(* IEC 61131-3 sources: plc-st-coding-agent/progress/evidence/full_r8_20261110b/native_evidence/codex_minimax-m27/public-easy-04/1, 1 file *)

(* ---- candidate.st ---- *)
FUNCTION_BLOCK FB
VAR_INPUT
    VISCOSITY_OK      : BOOL;
    PASTE_E_STOP_NC   : BOOL;
    DebounceMs        : DINT;
    CycleMs           : DINT;
END_VAR
VAR_OUTPUT
    VFD_RUN           : BOOL;
    PUMP_MAINT_DUE    : BOOL;
    PUMP_RUNTIME_ACC  : LINT;
END_VAR
VAR
    valid_duration     : DINT;
    prev_viscosity_ok  : BOOL;
    prev_paste_e_stop_nc : BOOL;
    prev_valid_duration : DINT;
    prev_vfd_run       : BOOL;
END_VAR

    IF NOT (PASTE_E_STOP_NC AND VISCOSITY_OK) THEN
        VFD_RUN := FALSE;
        valid_duration := 0;
    ELSE
        IF NOT prev_viscosity_ok OR NOT prev_paste_e_stop_nc THEN
            valid_duration := prev_valid_duration + CycleMs;
            VFD_RUN := (valid_duration >= DebounceMs);
        ELSIF prev_vfd_run THEN
            valid_duration := valid_duration + CycleMs;
            VFD_RUN := TRUE;
        ELSE
            valid_duration := valid_duration + CycleMs;
            VFD_RUN := (valid_duration >= DebounceMs);
        END_IF
    END_IF

    IF VFD_RUN THEN
        PUMP_RUNTIME_ACC := PUMP_RUNTIME_ACC + CycleMs;
    END_IF

    PUMP_MAINT_DUE := (PUMP_RUNTIME_ACC >= 1800000000);

    prev_valid_duration := valid_duration;
    prev_viscosity_ok := VISCOSITY_OK;
    prev_paste_e_stop_nc := PASTE_E_STOP_NC;
    prev_vfd_run := VFD_RUN;
END_FUNCTION_BLOCK
